// TIA Portal V21 export
// export: Created 2026-08-21T20:18:54.9081065Z, ExportSetting None, DisplayName Totally Integrated Automation Portal, DisplayVersion V21, DisplayName STEP 7 Professional, DisplayVersion V21, DisplayName STEP 7 Safety, DisplayVersion V21, DisplayName Tech WebApplication, DisplayVersion V21, DisplayName WinCC Basic/Comfort/Advanced, DisplayVersion V21, DisplayName WinCC Professional, DisplayVersion V21, DisplayName WinCC Unified, DisplayVersion V21
TYPE "UDT_MTP_BinProcessValueOut"
   STRUCT
      WQC { ExternalWritable := 'False'} : Byte := 16#FF;   // Worst Quality Code CCC
      V { ExternalWritable := 'False'} : Bool;   // External Source Value
      VState0 { ExternalWritable := 'False'} : String[16];   // Text Replacement Value (False)
      VState1 { ExternalWritable := 'False'} : String[16];   // Text Replacement Value (True)
   END_STRUCT;
END_TYPE
